(* IEC 61131-3 sources: SortJet_MasterSPS_Aufbau.fbsproj/07_Auftragsverwaltung/Job_Shuttle.prg.st^, 9 files *)

(* ---- Auftraege.act.st ---- *)
(* METADATA
{
	"v3Meta": {
		"objectGuid": "374beb49-ca7f-40e9-b2ab-7b5100759e7c"
	}
}
*)
ACTION Auftraege
//-------------------------------------------------------------------------------------------------
// AUFTRAG: M_SB0_MMI_SHEET_ORDER_SHUTTLE
//-------------------------------------------------------------------------------------------------
(* Hinweis:
   - Auftragsdaten an ein Shuttle uebergeben
*)
IF ( M_SB0_MMI_SHEET_ORDER_SHUTTLE ) THEN

  CASE tMmi2SpsInfo.wStationsNr OF

    cERSTES_SHUTTLE..cLETZTES_SHUTTLE:
      LocalAuftragsSpeicher REF= AuftragsSpeicherWand[tMmi2SpsInfo.wStationsNr, tMmi2SpsInfo.wAuftragsWand];
      M_SB0_MMI_SHEET_ORDER_SHUTTLE := FALSE;

    cERSTES_TRANSFERSHUTTLE..cLETZTES_TRANSFERSHUTTLE:
      LocalAuftragsSpeicher REF= AuftragsSpeicherTransfershuttle[tMmi2SpsInfo.wStationsNr];
      M_SB0_MMI_SHEET_ORDER_SHUTTLE := FALSE;

  END_CASE

  IF __ISVALIDREF(LocalAuftragsSpeicher) THEN

    LocalAuftragsSpeicher.NeuerAuftrag.wStationsNr            := tMmi2SpsInfo.wStationsNr;
    LocalAuftragsSpeicher.NeuerAuftrag.rVorabPosition         := tMmi2SpsInfo.rStationsPosition;
    LocalAuftragsSpeicher.NeuerAuftrag.rStationsZielposition  := tMmi2SpsInfo.rStationsPosition;     // Stationsposition der Quellstation
    LocalAuftragsSpeicher.NeuerAuftrag.rAuftragsLaenge        := tMmi2SpsInfo.rAuftragsLaenge;       // Länge der Scheibe/Batch
    LocalAuftragsSpeicher.NeuerAuftrag.rAuftragsHoehe         := tMmi2SpsInfo.rAuftragsHoehe;        // Höhe der Scheibe/Batch
    LocalAuftragsSpeicher.NeuerAuftrag.rAuftragsDicke         := tMmi2SpsInfo.rAuftragsDicke;        // Dicke der Scheibe/Batch
    LocalAuftragsSpeicher.NeuerAuftrag.wErsteLetzteScheibe    := tMmi2SpsInfo.wErsteLetzteScheibe;  // Kennzeichnung Erste und Letzte Scheibe
    LocalAuftragsSpeicher.NeuerAuftrag.wAnzahlScheiben        := tMmi2SpsInfo.wAnzahlScheiben;       // Anzahl der Scheiben
    LocalAuftragsSpeicher.NeuerAuftrag.wStationsWand          := tMmi2SpsInfo.wAuftragsWand;         // Stationswand der Quellstation
    LocalAuftragsSpeicher.NeuerAuftrag.wTransferstationsNr1   := tMmi2SpsInfo.wTransferstationsNr1;  // Stationsnummer der Zielstation 1
    LocalAuftragsSpeicher.NeuerAuftrag.wTransferstationsNr2   := tMmi2SpsInfo.wTransferstationsNr2;  // Stationsnummer der Zielstation 2
    LocalAuftragsSpeicher.NeuerAuftrag.rTransferposition1     := tMmi2SpsInfo.rTransferposition1;    // Stationsposition der Zielstation 1
    LocalAuftragsSpeicher.NeuerAuftrag.rTransferposition2     := tMmi2SpsInfo.rTransferposition2;    // Stationsposition der Zielstation 2
    LocalAuftragsSpeicher.NeuerAuftrag.wTransferwand          := tMmi2SpsInfo.wTransferwand;         // Stationswand der Zielstationen 1
    LocalAuftragsSpeicher.NeuerAuftrag.stAuftragsInformationen.wAuftragsInformationen := tMmi2SpsInfo.wAuftragsTyp;            // Zusaetzliche Auftrags- Informationen

    // Soll Drehpos der Folgestation für den Eintransport
    LocalAuftragsSpeicher.NeuerAuftrag.wTransferVersatzVorne   := tMmi2SpsInfo.rTransferstationModellversatzVorne;
    // Soll Drehpos der Folgestation nach dem Eintransport
    LocalAuftragsSpeicher.NeuerAuftrag.wTransferVersatzHinten  := tMmi2SpsInfo.rTransferstationModellversatzHinten;

    (* Hinweis:
       - Zuweisung der Bits "erste" und "letzte" Scheibe
    *)
    ErsteUndLetzteScheibeBits( wpErsteUndLetzteScheibe:= tMmi2SpsInfo.wErsteLetzteScheibe ,
                               wpLetzteScheibe => wlLetzteScheibe,
                               wpErsteScheibe  => wlErsteScheibe );

    LocalAuftragsSpeicher.NeuerAuftrag.bLetzteScheibe  := wlLetzteScheibe > 0;   // Stationsposition der Zielstation 2
    LocalAuftragsSpeicher.NeuerAuftrag.bErsteScheibe   := wlErsteScheibe  > 0;        // Stationswand der Zielstationen

    (* Hinweis:
       - 0 -> Eintransport
       - 1 -> Austransport
    *)
    IF ( tMmi2SpsInfo.wAuftragsTyp.0 ) THEN
      LocalAuftragsSpeicher.NeuerAuftrag.wAuftrag := eStation_Austransport;
    ELSE
      LocalAuftragsSpeicher.NeuerAuftrag.wAuftrag := eStation_Eintransport;
    END_IF

    LocalAuftragsSpeicher(bpNeuerAuftrag := TRUE);

  END_IF

END_IF

//-------------------------------------------------------------------------------------------------
// AUFTRAG: M_SB0_MMI_SortierungInsertExtractionShuttleData
//-------------------------------------------------------------------------------------------------
(* Hinweis:
   - Austransportschlitten mit einem Scheibenvortransport-Auftrag versehen
*)
IF ( M_SB0_MMI_SortierungInsertExtractionShuttleData ) THEN

  M_SB0_MMI_SortierungInsertExtractionShuttleData := FALSE;

  IF ( bgTransfershuttleVortransportAktivieren ) THEN

    // ---------------------------------------------------------------------------------------
    //  TRANSFERSHUTTLE VORTRANSPORT
    //
    //  Hinweis:
    //  - VortransportNummer_TS2 = 0   => Vortransport mit nur einem Transfershuttle
    //  - VortransportNummer_TS1 <> 0  => Vortransport im Transfershuttle-Verbund
    // ---------------------------------------------------------------------------------------
    IF ( tMmi2SpsInfo.wVortransportNummer_TS2 = 0  ) THEN

      AuftragsSpeicherTransfershuttle[tMmi2SpsInfo.wVortransportNummer_TS1].NeuerAuftrag.rStationsZielposition := tMmi2SpsInfo.rVortransportSollPosition_TS1;
      AuftragsSpeicherTransfershuttle[tMmi2SpsInfo.wVortransportNummer_TS1].NeuerAuftrag.rAuftragsLaenge       := tMmi2SpsInfo.rVortransportStrecke;
      AuftragsSpeicherTransfershuttle[tMmi2SpsInfo.wVortransportNummer_TS1].NeuerAuftrag.wTransferstationsNr1  := 0;
      AuftragsSpeicherTransfershuttle[tMmi2SpsInfo.wVortransportNummer_TS1].NeuerAuftrag.wTransferstationsNr2  := 0;
      AuftragsSpeicherTransfershuttle[tMmi2SpsInfo.wVortransportNummer_TS1].NeuerAuftrag.rTransferposition1    := tMmi2SpsInfo.rVortransportSollPosition_TS1;
      AuftragsSpeicherTransfershuttle[tMmi2SpsInfo.wVortransportNummer_TS1].NeuerAuftrag.rTransferposition2    := 0;
      AuftragsSpeicherTransfershuttle[tMmi2SpsInfo.wVortransportNummer_TS1].NeuerAuftrag.stAuftragsInformationen.cBIT_BUFFERSLOT_THICKNESS := ( tMmi2SpsInfo.wSlotThickness = 1 );
      AuftragsSpeicherTransfershuttle[tMmi2SpsInfo.wVortransportNummer_TS1].NeuerAuftrag.wAuftrag := eStation_Vortransport;
      AuftragsSpeicherTransfershuttle[tMmi2SpsInfo.wVortransportNummer_TS1](bpNeuerAuftrag := TRUE);

    ELSE
      VailiderenTransfershuttleVerbund ( wTransferstation1 := tMmi2SpsInfo.wVortransportNummer_TS1 ,
                                         wTransferstation2 := tMmi2SpsInfo.wVortransportNummer_TS2 ,
                                         wTransferstationMaster => tMmi2SpsInfo.wVortransportNummer_TS1,
                                         wTransferstationSlave  => tMmi2SpsInfo.wVortransportNummer_TS2 );

      AuftragsSpeicherTransfershuttle[tMmi2SpsInfo.wVortransportNummer_TS1].NeuerAuftrag.rStationsZielposition := tMmi2SpsInfo.rVortransportSollPosition_TS1;
      AuftragsSpeicherTransfershuttle[tMmi2SpsInfo.wVortransportNummer_TS1].NeuerAuftrag.rAuftragsLaenge       := tMmi2SpsInfo.rVortransportStrecke;
      AuftragsSpeicherTransfershuttle[tMmi2SpsInfo.wVortransportNummer_TS1].NeuerAuftrag.wTransferstationsNr1  := tMmi2SpsInfo.wVortransportNummer_TS1;
      AuftragsSpeicherTransfershuttle[tMmi2SpsInfo.wVortransportNummer_TS1].NeuerAuftrag.wTransferstationsNr2  := tMmi2SpsInfo.wVortransportNummer_TS2;
      AuftragsSpeicherTransfershuttle[tMmi2SpsInfo.wVortransportNummer_TS1].NeuerAuftrag.rTransferposition1    := tMmi2SpsInfo.rVortransportSollPosition_TS1;
      AuftragsSpeicherTransfershuttle[tMmi2SpsInfo.wVortransportNummer_TS1].NeuerAuftrag.rTransferposition2    := tMmi2SpsInfo.rVortransportSollPosition_TS2;
      AuftragsSpeicherTransfershuttle[tMmi2SpsInfo.wVortransportNummer_TS1].NeuerAuftrag.stAuftragsInformationen.cBIT_BUFFERSLOT_THICKNESS := ( tMmi2SpsInfo.wSlotThickness = 1 );
      AuftragsSpeicherTransfershuttle[tMmi2SpsInfo.wVortransportNummer_TS1].NeuerAuftrag.wAuftrag              := eStation_Vortransport;
      AuftragsSpeicherTransfershuttle[tMmi2SpsInfo.wVortransportNummer_TS1](bpNeuerAuftrag := TRUE);

    END_IF

  ELSE

    (* Hinweis:
       - Quittierung des Vortransportes
    *)
    wSps2MmiQuittierungVortransportStationsNr1 := tMmi2SpsInfo.wVortransportNummer_TS1;
    wSps2MmiQuittierungVortransportStationsNr2 := tMmi2SpsInfo.wVortransportNummer_TS2;
    wSps2MmiQuittierungVortransportStatus      := 1; // 0  = nicht Erfolgreich / 1 = erfolgreich
    rSps2MmiQuittierungVortransportWegStrecke  := tMmi2SpsInfo.rVortransportStrecke;

    MsgToMmi(auftragsnr_w := SB0_SPS_SortierungQuittExtractionShuttleData );

  END_IF

END_IF

//-------------------------------------------------------------------------------------------------
// AUFTRAG: M_SB0_MMI_SHUTTLE_INFORMATION
//-------------------------------------------------------------------------------------------------
IF ( M_SB0_MMI_SHUTTLE_INFORMATION ) THEN

  M_SB0_MMI_SHUTTLE_INFORMATION := FALSE;

  CASE tMmi2SpsInfo.wAuftrag_ShuttleNummer OF

    cERSTE_STATION..cLETZTE_STATION:
      ;
    cERSTES_SHUTTLE..cLETZTES_SHUTTLE:
      // Rueckfall: Schickt das MMI keine Wand (0), gilt Wand 1
      IF tMmi2SpsInfo.wAuftrag_ShuttleWand = 0 THEN
        tMmi2SpsInfo.wAuftrag_ShuttleWand := cWAND_1;
      END_IF
      CASE tMmi2SpsInfo.wAuftrag_ShuttleWand OF

          cWAND_1,
            cWAND_2:
          IF ( VorAbAuftragsDaten[tMmi2SpsInfo.wAuftrag_ShuttleNummer, tMmi2SpsInfo.wAuftrag_ShuttleWand].wAuftrag = eStation_Kein_Auftrag ) THEN
            VorAbAuftragsDaten[tMmi2SpsInfo.wAuftrag_ShuttleNummer, tMmi2SpsInfo.wAuftrag_ShuttleWand].rLaenge                := tMmi2SpsInfo.rAuftrag_Laenge;
            VorAbAuftragsDaten[tMmi2SpsInfo.wAuftrag_ShuttleNummer, tMmi2SpsInfo.wAuftrag_ShuttleWand].rDicke                 := tMmi2SpsInfo.rAuftrag_Dicke;
            VorAbAuftragsDaten[tMmi2SpsInfo.wAuftrag_ShuttleNummer, tMmi2SpsInfo.wAuftrag_ShuttleWand].wTransferStation       := tMmi2SpsInfo.wAuftrag_TranferStation;
            VorAbAuftragsDaten[tMmi2SpsInfo.wAuftrag_ShuttleNummer, tMmi2SpsInfo.wAuftrag_ShuttleWand].wAuftragstyp           := tMmi2SpsInfo.wAuftrag_Modus;
            VorAbAuftragsDaten[tMmi2SpsInfo.wAuftrag_ShuttleNummer, tMmi2SpsInfo.wAuftrag_ShuttleWand].wShuttleWandNummer     := tMmi2SpsInfo.wAuftrag_ShuttleWand;
            VorAbAuftragsDaten[tMmi2SpsInfo.wAuftrag_ShuttleNummer, tMmi2SpsInfo.wAuftrag_ShuttleWand].wTransferWand          := tMmi2SpsInfo.wAuftrag_TransferWand;
            VorAbAuftragsDaten[tMmi2SpsInfo.wAuftrag_ShuttleNummer, tMmi2SpsInfo.wAuftrag_ShuttleWand].wShuttleNummer         := tMmi2SpsInfo.wAuftrag_ShuttleNummer;

            VorAbAuftragsDaten[tMmi2SpsInfo.wAuftrag_ShuttleNummer, tMmi2SpsInfo.wAuftrag_ShuttleWand].stAuftragsInformationen.wAuftragsInformationen := tMmi2SpsInfo.wAuftrag_Modus;
            VorAbAuftragsDaten[tMmi2SpsInfo.wAuftrag_ShuttleNummer, tMmi2SpsInfo.wAuftrag_ShuttleWand].wAuftrag := eStation_VorabAuftrag;

          END_IF

        cWAND_1_2: //eigentlich Wand 1 und 2, da dies Bitcodiert ist, kommt dies als Wand3
          FOR wlIndexWand := cWAND_1 TO cANZAHL_WAENDE DO

            IF ( VorAbAuftragsDaten[tMmi2SpsInfo.wAuftrag_ShuttleNummer, wlIndexWand].wAuftrag = eStation_Kein_Auftrag ) THEN

              VorAbAuftragsDaten[tMmi2SpsInfo.wAuftrag_ShuttleNummer, wlIndexWand].rLaenge                := tMmi2SpsInfo.rAuftrag_Laenge;
              VorAbAuftragsDaten[tMmi2SpsInfo.wAuftrag_ShuttleNummer, wlIndexWand].rDicke                 := tMmi2SpsInfo.rAuftrag_Dicke;
              VorAbAuftragsDaten[tMmi2SpsInfo.wAuftrag_ShuttleNummer, wlIndexWand].wTransferStation       := tMmi2SpsInfo.wAuftrag_TranferStation;
              VorAbAuftragsDaten[tMmi2SpsInfo.wAuftrag_ShuttleNummer, wlIndexWand].wAuftragstyp           := tMmi2SpsInfo.wAuftrag_Modus;
              VorAbAuftragsDaten[tMmi2SpsInfo.wAuftrag_ShuttleNummer, wlIndexWand].wShuttleWandNummer     := wlIndexWand;
              VorAbAuftragsDaten[tMmi2SpsInfo.wAuftrag_ShuttleNummer, wlIndexWand].wTransferWand          := tMmi2SpsInfo.wAuftrag_TransferWand;
              VorAbAuftragsDaten[tMmi2SpsInfo.wAuftrag_ShuttleNummer, wlIndexWand].wShuttleNummer         := tMmi2SpsInfo.wAuftrag_ShuttleNummer;

              VorAbAuftragsDaten[tMmi2SpsInfo.wAuftrag_ShuttleNummer, wlIndexWand].stAuftragsInformationen.wAuftragsInformationen := tMmi2SpsInfo.wAuftrag_Modus;
              VorAbAuftragsDaten[tMmi2SpsInfo.wAuftrag_ShuttleNummer, wlIndexWand].wAuftrag := eStation_VorabAuftrag;

            END_IF

          END_FOR

        ELSE
          ;

      END_CASE

    cERSTES_TRANSFERSHUTTLE..cLETZTES_TRANSFERSHUTTLE:
      IF ( NOT Job_Shuttle.abpStarteParalleleBausteinAnsteuerung[tMmi2SpsInfo.wAuftrag_ShuttleNummer] ) THEN
        Job_Shuttle.VorAbAuftragsDaten[tMmi2SpsInfo.wAuftrag_ShuttleNummer, cWAND_1].rLaenge                := tMmi2SpsInfo.rAuftrag_Laenge;
        Job_Shuttle.VorAbAuftragsDaten[tMmi2SpsInfo.wAuftrag_ShuttleNummer, cWAND_1].rDicke                 := tMmi2SpsInfo.rAuftrag_Dicke;
        Job_Shuttle.VorAbAuftragsDaten[tMmi2SpsInfo.wAuftrag_ShuttleNummer, cWAND_1].wTransferStation       := tMmi2SpsInfo.wAuftrag_TranferStation;
        Job_Shuttle.VorAbAuftragsDaten[tMmi2SpsInfo.wAuftrag_ShuttleNummer, cWAND_1].wAuftragstyp           := tMmi2SpsInfo.wAuftrag_Modus;
        Job_Shuttle.VorAbAuftragsDaten[tMmi2SpsInfo.wAuftrag_ShuttleNummer, cWAND_1].wShuttleWandNummer     := tMmi2SpsInfo.wAuftrag_ShuttleWand;
        Job_Shuttle.VorAbAuftragsDaten[tMmi2SpsInfo.wAuftrag_ShuttleNummer, cWAND_1].wTransferWand          := tMmi2SpsInfo.wAuftrag_TransferWand;
        Job_Shuttle.VorAbAuftragsDaten[tMmi2SpsInfo.wAuftrag_ShuttleNummer, cWAND_1].wShuttleNummer         := tMmi2SpsInfo.wAuftrag_ShuttleNummer;

        Job_Shuttle.VorAbAuftragsDaten[tMmi2SpsInfo.wAuftrag_ShuttleNummer, cWAND_1].stAuftragsInformationen.wAuftragsInformationen := tMmi2SpsInfo.wAuftrag_Modus;

        Job_Shuttle.abpStarteParalleleBausteinAnsteuerung[tMmi2SpsInfo.wAuftrag_ShuttleNummer] := TRUE;
      END_IF

    ELSE
      (* Fehlerbehandlung:
      *)
      wpgFehlerdaten[0] := tMmi2SpsInfo.wAuftrag_ShuttleNummer;
      wpgFehlerdaten[1] := tMmi2SpsInfo.wAuftrag_TranferStation;
      SpsError( eFehler_Station,
                cMELDUNG_AUFTRAGSDATEN_UNGUELTIGE_STATION,
                tMmi2SpsInfo.wAuftrag_ShuttleNummer,
                AutomatikkreisBestimmen(tMmi2SpsInfo.wAuftrag_ShuttleNummer),
                wpgFehlerdaten );

  END_CASE

END_IF

//-------------------------------------------------------------------------------------------------
// AUFTRAG: M_SB0_MMI_GETSORTIERUNGSHUTTLEPOS
//-------------------------------------------------------------------------------------------------
(* Hinweis:
   - Verfarhlogik
     => Absetzen der Positionen
     => Melden der IST- Position wenn die Positionierung aufgrund eines
        Fehler [ Verfahrfreigabe fehlt ] nicht durchgefuehrt werden kann
*)
IF ( M_SB0_MMI_GETSORTIERUNGSHUTTLEPOS ) THEN

  M_SB0_MMI_GETSORTIERUNGSHUTTLEPOS := FALSE;

  SendShuttlePosition();

END_IF

//-------------------------------------------------------------------------------------------------
// AUFTRAG: M_SB0_MMI_TS_REPOSITIONING_LITES
//-------------------------------------------------------------------------------------------------

(* Hinweis:
   - Funktion zum zurueckfahren der Glaeser und neu Positionieren im Speicher
*)
IF ( M_SB0_MMI_TS_REPOSITIONING_LITES ) THEN
  M_SB0_MMI_TS_REPOSITIONING_LITES := FALSE;

  CASE tMmi2SpsInfo.wStationsNr OF

    cERSTES_TRANSFERSHUTTLE..cLETZTES_TRANSFERSHUTTLE:
      AuftragsSpeicherTransfershuttle[tMmi2SpsInfo.wStationsNr].NeuerAuftrag.wStationsNr           := tMmi2SpsInfo.wStationsNr;
      AuftragsSpeicherTransfershuttle[tMmi2SpsInfo.wStationsNr].NeuerAuftrag.rStationsZielposition := tMmi2SpsInfo.rStationsPosition;
      AuftragsSpeicherTransfershuttle[tMmi2SpsInfo.wStationsNr].NeuerAuftrag.wTransferstationsNr1  := tMmi2SpsInfo.wTransferstationsNr1;
      AuftragsSpeicherTransfershuttle[tMmi2SpsInfo.wStationsNr].NeuerAuftrag.rModellVersatzHinten  := tMmi2SpsInfo.rModellversatzHinten;

      IF ( tMmi2SpsInfo.rAuftragsDicke = 0 ) THEN
        AuftragsSpeicherTransfershuttle[tMmi2SpsInfo.wStationsNr].NeuerAuftrag.rAuftragsDicke        := 4.0;
      ELSE
        AuftragsSpeicherTransfershuttle[tMmi2SpsInfo.wStationsNr].NeuerAuftrag.rAuftragsDicke        := 19.0;
      END_IF

      AuftragsSpeicherTransfershuttle[tMmi2SpsInfo.wStationsNr].NeuerAuftrag.wAuftrag := eStation_Scheibenkorrektur;
      AuftragsSpeicherTransfershuttle[tMmi2SpsInfo.wStationsNr](bpNeuerAuftrag := TRUE);

      AuftragsSpeicherTransfershuttle[tMmi2SpsInfo.wTransferstationsNr1].NeuerAuftrag.wStationsNr           := tMmi2SpsInfo.wTransferstationsNr1;
      AuftragsSpeicherTransfershuttle[tMmi2SpsInfo.wTransferstationsNr1].NeuerAuftrag.rStationsZielposition := tMmi2SpsInfo.rTransferposition1;
      AuftragsSpeicherTransfershuttle[tMmi2SpsInfo.wTransferstationsNr1].NeuerAuftrag.wTransferstationsNr1  := tMmi2SpsInfo.wStationsNr;
      AuftragsSpeicherTransfershuttle[tMmi2SpsInfo.wTransferstationsNr1].NeuerAuftrag.rModellVersatzHinten  := tMmi2SpsInfo.rModellversatzHinten;

      IF ( tMmi2SpsInfo.rAuftragsDicke = 0 ) THEN
        AuftragsSpeicherTransfershuttle[tMmi2SpsInfo.wTransferstationsNr1].NeuerAuftrag.rAuftragsDicke        := 4.0;
      ELSE
        AuftragsSpeicherTransfershuttle[tMmi2SpsInfo.wTransferstationsNr1].NeuerAuftrag.rAuftragsDicke        := 19.0;
      END_IF

      AuftragsSpeicherTransfershuttle[tMmi2SpsInfo.wTransferstationsNr1].NeuerAuftrag.wAuftrag := eStation_Transportkopplung;
      AuftragsSpeicherTransfershuttle[tMmi2SpsInfo.wTransferstationsNr1](bpNeuerAuftrag := TRUE);

  END_CASE

END_IF

//-------------------------------------------------------------------------------------------------
// AUFTRAG: M_SB0_MMI_SORTIERUNGCANcELSHUTTLEDATA
//-------------------------------------------------------------------------------------------------
(* Hinweis:
   - Abbrechen eines aktiven Shuttleauftrags
*)
IF ( M_SB0_MMI_SORTIERUNGCANCELSHUTTLEDATA ) THEN

  M_SB0_MMI_SortierungCancelShuttleData := FALSE;

  CASE tMmi2SpsInfo.wCancelShuttleDataShuttleNr OF

    cERSTES_SHUTTLE..cLETZTES_SHUTTLE:
      IF ( AuftragsdatenWand[tMmi2SpsInfo.wCancelShuttleDataShuttleNr, cWAND_1].wAuftrag <> eStation_Kein_Auftrag ) THEN
        AuftragsdatenWand[tMmi2SpsInfo.wCancelShuttleDataShuttleNr, cWAND_1].wAuftrag :=  eStation_Kein_Auftrag;
      END_IF

    cERSTES_TRANSFERSHUTTLE..cLETZTES_TRANSFERSHUTTLE:
      IF ( Job_Shuttle.AuftragsdatenTransfershuttle[tMmi2SpsInfo.wCancelShuttleDataShuttleNr].wAuftrag <> eStation_Kein_Auftrag ) THEN
        Job_Shuttle.AuftragsdatenTransfershuttle[tMmi2SpsInfo.wCancelShuttleDataShuttleNr].wAuftrag :=  eStation_Kein_Auftrag;
      END_IF

  END_CASE

END_IF

//-------------------------------------------------------------------------------------------------
// S T A R T - Fächerwagen Suche mittels Sensor
//-------------------------------------------------------------------------------------------------

IF ( M_SB0_MMI_POSITIONMEASUREONOFF ) THEN

  M_SB0_MMI_POSITIONMEASUREONOFF := FALSE;

  IF ( tMmi2SpsInfo.wShuttleFWSucheAN_AUS = 1 ) THEN
    AuftragsSpeicherWand[tMmi2SpsInfo.wShuttleNummerFWSuche, cWAND_1].NeuerAuftrag.wAuftrag := eStation_RackSuche;
    AuftragsSpeicherWand[tMmi2SpsInfo.wShuttleNummerFWSuche, cWAND_1](bpNeuerAuftrag := TRUE);
  ELSE
    IF ( AuftragsdatenWand[tMmi2SpsInfo.wShuttleNummerFWSuche, cWAND_1].wAuftrag = eStation_RackSuche ) THEN
      AuftragsdatenWand[tMmi2SpsInfo.wShuttleNummerFWSuche, cWAND_1].wAuftrag := eStation_Kein_Auftrag;
    END_IF
  END_IF

END_IF

//-------------------------------------------------------------------------------------------------
// SHUTTLE DEAKTIVIEREN VIA MMI
//-------------------------------------------------------------------------------------------------
IF ( M_SB0_MMI_STATIONSTATUS ) THEN

  CASE tMmi2SpsInfo.wStationsNummer OF

    cERSTES_SHUTTLE..cLETZTES_SHUTTLE:
      starrShuttleBasisParameter[tMmi2SpsInfo.wStationsNummer].stMKs.bDeaktivieren := tMmi2SpsInfo.wStationsStatusWord2.0;
      M_SB0_MMI_STATIONSTATUS := FALSE;

    cERSTES_TRANSFERSHUTTLE..cLETZTES_TRANSFERSHUTTLE:
      starrTransfershuttleBasisParameter[tMmi2SpsInfo.wStationsNummer].stMKs.bDeaktivieren := tMmi2SpsInfo.wStationsStatusWord2.0;
      M_SB0_MMI_STATIONSTATUS := FALSE;

  END_CASE

END_IF
END_ACTION

(* ---- Master_Transfershuttle.meth.st ---- *)
(* METADATA
{
	"v3Meta": {
		"objectGuid": "5a2b5255-704a-40f5-acbe-9caa573edc30"
	}
}
*)
METHOD INTERNAL Master_Transfershuttle
VAR_INPUT
  wStation : WORD;
END_VAR

// ****************************************************9*********************************************
// STEUERUNG: EINTRANSPORT
// *************************************************************************************************

IF ( AuftragsdatenTransfershuttle[wStation].wAuftrag = eStation_Eintransport ) THEN
  (* Hinweis:
     - Aufruf der Schrittkette
  *)
  TS_Eintransport[wStation]( Auftragsdaten := AuftragsdatenTransfershuttle[wStation], wStation := wStation );
  (* Hinweis:
     - Abschluss der Schrittkette
  *)
  IF TS_Eintransport[wStation].bpDone THEN
    AuftragsdatenTransfershuttle[wStation] := TS_Eintransport[wStation].Auftragsdaten;
    TS_Eintransport[wStation](bpReset := TRUE);
  END_IF
  (* Hinweis:
     - Fehler-Auswertung
  *)
  blFehlerTS[wStation] := TS_Eintransport[wStation].bpFehler;
  IF rtlFehlerTS[wStation].Q THEN
    IF ( starrTransfershuttleBasisParameter[wStation].bRueckwaertsTransportieren[cWAND_1] ) THEN
      AutomatikFehlerTransfershuttleSetzen(starrTransferShuttleBasisParameter[wStation].stMKs.eaAutomatikkreis, abpFehler, cSPEICHER_AUSLAUFSEITE);
      IF aTransfershuttles[wStation].bpAnforderungBetriebsstopp THEN
        AutomatikFehlerTransfershuttleSetzen(starrTransferShuttleBasisParameter[wStation].stMKs.eaAutomatikkreis, abpFehler, cSPEICHER_EINLAUFSEITE);
      END_IF
    ELSE
      AutomatikFehlerTransfershuttleSetzen(starrTransferShuttleBasisParameter[wStation].stMKs.eaAutomatikkreis, abpFehler, cSPEICHER_EINLAUFSEITE);
      IF aTransfershuttles[wStation].bpAnforderungBetriebsstopp THEN
        AutomatikFehlerTransfershuttleSetzen(starrTransferShuttleBasisParameter[wStation].stMKs.eaAutomatikkreis, abpFehler, cSPEICHER_AUSLAUFSEITE);
      END_IF
    END_IF
  END_IF
ELSE
  (* Hinweis:
     - Reset der Schrittkette
  *)
  IF ( TS_Eintransport[wStation].steplSchritt <> STEP_0_E ) THEN
    TS_Eintransport[wStation](bpReset := TRUE);
  END_IF
END_IF

// ****************************************************9*********************************************
// STEUERUNG: AUSTRANSPORT
// *************************************************************************************************

IF ( AuftragsdatenTransfershuttle[wStation].wAuftrag = eStation_Austransport ) THEN
  (* Hinweis:
     - Aufruf der Schrittkette
  *)
  TS_Austransport[wStation]( Auftragsdaten := AuftragsdatenTransfershuttle[wStation], wStation := wStation );
  (* Hinweis:
     - Abschluss der Schrittkette
  *)
  IF TS_Austransport[wStation].bpDone THEN
    AuftragsdatenTransfershuttle[wStation] := TS_Austransport[wStation].Auftragsdaten;
    TS_Austransport[wStation](bpReset := TRUE);
  END_IF
  (* Hinweis:
     - Fehler-Auswertung
  *)
  blFehlerTS[wStation] := TS_Austransport[wStation].bpFehler;
  IF rtlFehlerTS[wStation].Q THEN
    IF ( starrTransfershuttleBasisParameter[wStation].bRueckwaertsTransportieren[cWAND_1] ) THEN
      AutomatikFehlerTransfershuttleSetzen(starrTransferShuttleBasisParameter[wStation].stMKs.eaAutomatikkreis, abpFehler, cSPEICHER_EINLAUFSEITE);
      IF aTransfershuttles[wStation].bpAnforderungBetriebsstopp THEN
        AutomatikFehlerTransfershuttleSetzen(starrTransferShuttleBasisParameter[wStation].stMKs.eaAutomatikkreis, abpFehler, cSPEICHER_AUSLAUFSEITE);
      END_IF
    ELSE
      AutomatikFehlerTransfershuttleSetzen(starrTransferShuttleBasisParameter[wStation].stMKs.eaAutomatikkreis, abpFehler, cSPEICHER_AUSLAUFSEITE);
      IF aTransfershuttles[wStation].bpAnforderungBetriebsstopp THEN
        AutomatikFehlerTransfershuttleSetzen(starrTransferShuttleBasisParameter[wStation].stMKs.eaAutomatikkreis, abpFehler, cSPEICHER_EINLAUFSEITE);
      END_IF
    END_IF
  END_IF
ELSE
  (* Hinweis:
     - Reset der Schrittkette
  *)
  IF ( TS_Austransport[wStation].steplSchritt <> STEP_0_E ) THEN
    TS_Austransport[wStation](bpReset := TRUE);
  END_IF
END_IF

// ****************************************************9*********************************************
// STEUERUNG: VORTRANSPORT
// *************************************************************************************************

IF ( AuftragsdatenTransfershuttle[wStation].wAuftrag = eStation_Vortransport ) THEN
  (* Hinweis:
     - Aufruf der Schrittkette
  *)
  TS_Vortransport[wStation]( Auftragsdaten := AuftragsdatenTransfershuttle[wStation], wStation := wStation);
  (* Hinweis:
     - Abschluss der Schrittkette
  *)
  IF TS_Vortransport[wStation].bpDone THEN
    AuftragsdatenTransfershuttle[wStation] := TS_Vortransport[wStation].Auftragsdaten;
    TS_Vortransport[wStation](bpReset := TRUE);
  END_IF
  (* Hinweis:
     - Fehler-Auswertung
  *)
  blFehlerTS[wStation] := TS_Vortransport[wStation].bpFehler;
  IF rtlFehlerTS[wStation].Q THEN
    AutomatikFehlerSetzen(starrTransferShuttleBasisParameter[wStation].stMKs.eaAutomatikkreis, abpFehler);
  END_IF
ELSE
  (* Hinweis:
     - Reset der Schrittkette
  *)
  IF ( TS_Vortransport[wStation].steplSchritt <> STEP_0_E ) THEN
    TS_Vortransport[wStation](bpReset := TRUE);
  END_IF
END_IF

// ****************************************************9*********************************************
// STEUERUNG: QUERFAHRT
// *************************************************************************************************

IF ( AuftragsdatenTransfershuttle[wStation].wAuftrag = eStation_Vorabpositionierung ) THEN
  (* Hinweis:
     - Aufruf der Schrittkette
  *)
  TS_Querfahrt[wStation]( Auftragsdaten := AuftragsdatenTransfershuttle[wStation], wStation := wStation );
  (* Hinweis:
     - Abschluss der Schrittkette
  *)
  IF TS_Querfahrt[wStation].bpDone THEN
    AuftragsdatenTransfershuttle[wStation] := TS_Querfahrt[wStation].Auftragsdaten;
    TS_Querfahrt[wStation](bpReset := TRUE);
  END_IF
  (* Hinweis:
     - Fehler-Auswertung
  *)
  blFehlerTS[wStation] := TS_Querfahrt[wStation].bpFehler;
  IF rtlFehlerTS[wStation].Q THEN
    AutomatikFehlerSetzen(starrTransferShuttleBasisParameter[wStation].stMKs.eaAutomatikkreis, abpFehler);
  END_IF
ELSE
  (* Hinweis:
     - Reset der Schrittkette
  *)
  IF ( TS_Querfahrt[wStation].steplSchritt <> STEP_0_E ) THEN
    TS_Querfahrt[wStation](bpReset := TRUE);
  END_IF
END_IF

//-------------------------------------------------------------------------------------------------
// STEUERUNG: SPEICHERFACHVALIDIERUNG
//-------------------------------------------------------------------------------------------------
IF (  abpSpeicherfachValidierung[wStation] ) THEN
  CASE asteplSpeicherfachValidierung[wStation] OF
    // SPEICHERFACHVALIDIERUNG =============================
    STEP_0_E:
      (* Hinweis:
         - Option: Sicherstellen das der Output-Sicherheitskreis geschlossen ist
      *)
      IF checkSafetyCircuitsNotBlocked(starrTransferShuttleBasisParameter[wStation])
         AND NOT starrTransfershuttleBasisParameter[wStation].bReset
      THEN
        awlStatusSpeichervalidierung[wStation]   := cAUFTRAG_KEIN_STATUS;
        asteplSpeicherfachValidierung[wStation] := STEP_10_E;
      END_IF

    // SPEICHERFACHVALIDIERUNG =============================
    STEP_10_E:
      // ---------------------------------------------------------------------------------------
      //  PRUEFEN TRANSFERSHUTTLE VERBUND
      //
      //  Hinweis:
      //  - wTransfershuttle_Nummer2 = 0   => Vortransport mit nur einem Transfershuttle
      //  - wTransfershuttle_Nummer2 <> 0  => Vortransport im Transfershuttle-Verbund
      // ---------------------------------------------------------------------------------------

      IF ( starrAuftragsdatenSpeicherfachValidierung[wStation].wTransferstationsNr2 <> 0 )  THEN

        awlVerbundTransfershuttle[wStation] := AuftragsdatenTransfershuttle[wStation].wTransferstationsNr2;

        IF ( AuftragsdatenTransfershuttle[awlVerbundTransfershuttle[wStation]].wAuftrag = eStation_Kein_Auftrag ) THEN
          asteplSpeicherfachValidierung[wStation] := STEP_20_E;
        END_IF

      ELSE
        (* Hinweis:
           - Informationen uebergeben und die Validierung starten
        *)
        starrTransfershuttleBasisParameter[wStation].pAuftrag[cWAND_1] := starrAuftragsdatenSpeicherfachValidierung[wStation];
        aTransfershuttles[wStation].bpStarteSpeicherfachValidierung := TRUE;

        asteplSpeicherfachValidierung[wStation] := STEP_100_E;

      END_IF

    // SPEICHERFACHVALIDIERUNG =============================
    STEP_20_E:

      (* Hinweis:
         - Transfershuttle koppeln
      *)
      aTransfershuttles[wStation].stpInTransportVerbund                             := aTransfershuttles[awlVerbundTransfershuttle[wStation]].stpOutTransportVerbund;
      aTransfershuttles[awlVerbundTransfershuttle[wStation]].stpInTransportVerbund  := aTransfershuttles[wStation].stpOutTransportVerbund;

      (* Hinweis:
         - Auftragsdaten uebergeben
      *)
      AuftragsdatenTransfershuttle[awlVerbundTransfershuttle[wStation]].rAuftragsDicke        := starrAuftragsdatenSpeicherfachValidierung[wStation].rAuftragsDicke ;
      AuftragsdatenTransfershuttle[awlVerbundTransfershuttle[wStation]].rStationsZielposition := starrAuftragsdatenSpeicherfachValidierung[wStation].rTransferposition2 ;
      AuftragsdatenTransfershuttle[awlVerbundTransfershuttle[wStation]].wStationsNr           := starrAuftragsdatenSpeicherfachValidierung[wStation].wTransferstationsNr2 ;
      AuftragsdatenTransfershuttle[awlVerbundTransfershuttle[wStation]].wAuftrag              := eStation_Transportkopplung;

      (* Hinweis:
         - Auftragsdaten uebergeben
      *)
      starrTransfershuttleBasisParameter[wStation].pAuftrag[cWAND_1] := starrAuftragsdatenSpeicherfachValidierung[wStation];
      aTransfershuttles[wStation].bpStarteSpeicherfachValidierung := TRUE;

      asteplSpeicherfachValidierung[wStation] := STEP_100_E;

    // SPEICHERFACHVALIDIERUNG =============================
    STEP_100_E:
      // ---------------------------------------------------------------------------------------
      //  AUSWERTUNG TRANSFERSHUTTLE - SPEICHERFACH VALIDIERUNG
      //
      //  Hinweis:
      //  - n/c
      // ---------------------------------------------------------------------------------------

      IF ( aTransfershuttles[wStation].bpSpeicherfachValidierungAbgeschlossen ) THEN
        aTransfershuttles[wStation].bpStarteSpeicherfachValidierung := FALSE;
        awlStatusSpeichervalidierung[wStation] := cAUFTRAG_ERFOLGREICH;

        asteplSpeicherfachValidierung[wStation] := STEP_120_E;
      END_IF

      // Fehlverhalten
      IF ( starrTransfershuttleBasisParameter[wStation].bFehler ) THEN

        aTransfershuttles[wStation].bpStarteSpeicherfachValidierung := FALSE;
        awlStatusSpeichervalidierung[wStation] := cAUFTRAG_FEHLER;

        asteplSpeicherfachValidierung[wStation] := STEP_120_E;

        (* Hinweis:
           - Meldung an die HMI generieren.
             => Gesendet wird: Shuttlenummer \Position \Fehlertyp
        *)
        wgSps2MmiShuttleNr                 := starrTransfershuttleBasisParameter[wStation].stMKs.stStationsNummern.NummerIntern;
        rgSPS2MMIExtractionShuttlePosition := starrTransfershuttleBasisParameter[wStation].rAktuellePositionQuerfahrt;
        wSps2MmiFehlertyp                  := aTransfershuttles[wStation].wpAusnahmefehlerTyp;
        MsgToMmi(auftragsnr_w := SB0_SPS_TRANSFERSHUTTLEFEHLER );// Fehlermeldung ans MMI für den folgenden Systemcheck

        (* Hinweis:
           - Fehlermeldung generieren
        *)
        SpsError( eFehler_Station,
                  starrTransfershuttleBasisParameter[wStation].wFehlerNummer,
                  starrTransfershuttleBasisParameter[wStation].stMKs.stStationsNummern.NummerIntern,
                  AutomatikkreisBestimmen(starrTransfershuttleBasisParameter[wStation].stMKs.stStationsNummern.NummerSPS),
                  starrTransfershuttleBasisParameter[wStation].awFehlerInformationen );

      END_IF

    // SPEICHERFACHVALIDIERUNG =============================
    STEP_120_E:
      wgSps2MmiShuttleNr         := starrTransfershuttleBasisParameter[wStation].stMKs.stStationsNummern.NummerIntern;
      wSps2MmiValidierungsStatus := awlStatusSpeichervalidierung[wStation];
      MsgToMmi(auftragsnr_w := SB0_SPS_TRANSFERSHUTTLECHECK_ABGESCHLOSSEN );// Fehlermeldung ans MMI für den folgenden Systemcheck

      asteplSpeicherfachValidierung[wStation] := SEL( awlStatusSpeichervalidierung[wStation] = cAUFTRAG_FEHLER,
                                                      STEP_1000_E,
                                                      STEP_900_E );

    // SPEICHERFACHVALIDIERUNG =============================
    STEP_900_E:
      AutomatikFehlerSetzen(starrTransferShuttleBasisParameter[wStation].stMKs.eaAutomatikkreis, abpFehler);

    // SPEICHERFACHVALIDIERUNG =============================
    STEP_1000_E:
      abpSpeicherfachValidierung[wStation] := FALSE;

      (* Hinweis:
         - Pruefen ob die Transferkopplung geloest werden muss
      *)
      IF ( PruefungWertImIntervall(AuftragsdatenTransfershuttle[wStation].wTransferstationsNr2, cERSTES_TRANSFERSHUTTLE, cLETZTES_TRANSFERSHUTTLE) ) THEN

        IF ( AuftragsdatenTransfershuttle[AuftragsdatenTransfershuttle[wStation].wTransferstationsNr2].wAuftrag = eStation_Transportkopplung ) THEN
          AuftragsdatenTransfershuttle[AuftragsdatenTransfershuttle[wStation].wTransferstationsNr2].wAuftrag := eStation_Kein_Auftrag;
        END_IF

      END_IF

  // SPEICHERFACHVALIDIERUNG =============================
  END_CASE

END_IF

IF ( NOT abpSpeicherfachValidierung[wStation] ) THEN

  IF ( asteplSpeicherfachValidierung[wStation] > STEP_0_E ) THEN
    aTransfershuttles[wStation].bpStarteSpeicherfachValidierung := FALSE;
    asteplSpeicherfachValidierung[wStation] := STEP_0_E;
  END_IF

END_IF
END_METHOD

(* ---- Meldungen.act.st ---- *)
(* METADATA
{
	"v3Meta": {
		"objectGuid": "68e675d5-67ba-4597-82c1-c0511fb282bc"
	}
}
*)
ACTION Meldungen
//-------------------------------------------------------------------------------------------------
// AKTION: MELDUNGEN
//-------------------------------------------------------------------------------------------------
// WatchIO:
//   - Ueberwachung der Verfahrfreigabe der Shuttle
//     -> Inputshuttle
//     -> Outputshuttle
//     -> Transfershuttle
FOR wlIndex := cERSTES_SHUTTLE TO cLETZTES_SHUTTLE DO
  WatchIo( NOT abgVerfahrfreigabeShuttle[wlIndex], ioccShuttle1VerfahrfreigabeFehlt + (wlIndex - 101) );
END_FOR;

FOR wlIndex := cERSTES_TRANSFERSHUTTLE TO cLETZTES_TRANSFERSHUTTLE DO
  WatchIo( NOT abgVerfahrfreigabeShuttle[wlIndex], ioccTransfershuttle1VerfahrfreigabeFehlt + (wlIndex - 151) );
END_FOR;
END_ACTION

(* ---- Reset.act.st ---- *)
(* METADATA
{
	"v3Meta": {
		"objectGuid": "238ec719-f16e-4d9c-9f71-7a8241f71645"
	}
}
*)
ACTION Reset
//-------------------------------------------------------------------------------------------------
// AKTION: RESET
//-------------------------------------------------------------------------------------------------

(* Hinweis:
   - Zuruecksetzen des AK
     => Inputshuttle [expliziet]
*)
FOR wlIndexReset := cERSTER_AUTOMATIKKREIS TO cLETZTER_AUTOMATIKKREIS DO

  IF abpReset[wlIndexReset] THEN

    abpReset[wlIndexReset] := FALSE;
    abpFehler[wlIndexReset] := FALSE;

    FOR wlIndex := cERSTES_SHUTTLE TO cLETZTES_SHUTTLE DO
      IF StationInAutomatikkreis(starrShuttleBasisParameter[wlIndex].stMKs.eaAutomatikkreis, wlIndexReset) THEN
        AuftragsSpeicherShuttle[wlIndex].bpReset := TRUE;
        AuftragsSpeicherShuttle[wlIndex]();

        abgVerfahrfreigabeShuttle[wlindex] := TRUE;

        AuftragsdatenStation[wlIndex].wAuftrag := eStation_Kein_Auftrag;

        starrShuttleBasisParameter[wlIndex].bReset := TRUE;

        Querfahrt[wlIndex]( bpReset := TRUE );
        Racksuche[wlIndex]( bpReset := TRUE );

        FOR wlIndexWand := cWAND_1 TO cANZAHL_WAENDE DO

          AuftragsSpeicherWand[wlIndex,wlIndexWand].bpReset := TRUE;
          AuftragsSpeicherWand[wlIndex,wlIndexWand]();

          Eintransport[wlIndex, wlIndexWand]( bpReset := TRUE );
          Austransport[wlIndex, wlIndexWand]( bpReset := TRUE );

          VorabkomponentenAnsteuerung[wlIndex, wlIndexWand]( bpReset := TRUE );

          AuftragsdatenWand[wlIndex, wlIndexWand].wAuftrag := eStation_Kein_Auftrag;
          VorAbAuftragsDaten[wlIndex, wlIndexWand].wAuftrag := eStation_Kein_Auftrag;

          blFehler[wlIndex, wlIndexWand] := FALSE;

          starrShuttleBasisParameter[wlIndex].bEintransportGewesen[wlIndexWand] := FALSE;
        END_FOR

      END_IF
    END_FOR

    FOR wlIndex := cERSTES_TRANSFERSHUTTLE TO cLETZTES_TRANSFERSHUTTLE  DO

      // WICHTIG: OR_ELSE -> ZWEITE BEDINGUNG WIRD NUR GEPRÜFT, WENN ERSTE FALSE IST !!! IST DIE ERSTE FALSE, WIRD DIE 2. BEDINGUNG GEPRÜFT ; IST DIE ERSTE TRUE, WIRD DIE 2. BEDINGUNG IGNORIERT UND NICHT MEHR GEPRÜFT (wg. ZUGRIFFSVERLETZTUNG)
      // Alle konfigurierten Automatikkreise des TS sind in Hand
      // ODER
      // Output-AK ist nicht in den vorhandenen Automatikkreisen der Maschine definiert ; das heißt, Erster AK = 1 und ANZAHL < wlAutomatikkreis2 --- OR_ELSE der 2. konfigurierte Automatikkreis für das TS ist 0; somit ist das TS nur in einem AK definiert
      IF   ( NOT AutomatikAktiv(wlIndex)
             OR ( ( cANZAHL_AUTOMATIKKREISE = 1 ) OR_ELSE ( starrTransfershuttleBasisParameter[wlIndex].stMKs.eaAutomatikkreis[wlAutomatikkreis2] = 0 ) ) )
           AND StationInAutomatikkreis(starrTransfershuttleBasisParameter[wlIndex].stMKs.eaAutomatikkreis, wlIndexReset)
      THEN
        AuftragsSpeicherTransfershuttle[wlIndex].bpReset := TRUE;
        AuftragsSpeicherTransfershuttle[wlIndex]();

        abgVerfahrfreigabeShuttle[wlindex] := TRUE;

        abpStarteParalleleBausteinAnsteuerung[wlIndex] := FALSE;
        abpSpeicherfachValidierung[wlIndex]  := FALSE;
        AuftragsdatenTransfershuttle[wlIndex].wAuftrag := eStation_Kein_Auftrag;
        starrTransferShuttleBasisParameter[wlIndex].bReset := TRUE;
        blFehlerTS[wlIndex] := FALSE;

      ELSE

        // Der zu resettende AK entspricht dem ERSTEN (INPUTSEITE) konfigurierten AK des TS
        // UND Doppelte Sicherheit: Nochmal prüfen, dass das TS im zu resetten AK ist
        // UND Automatik des zu resettenden AK darf NICHT mehr TRUE sein
        IF                ( wlIndexReset = starrTransfershuttleBasisParameter[wlIndex].stMKs.eaAutomatikkreis[1] )
                 AND_THEN StationInAutomatikkreis(starrTransfershuttleBasisParameter[wlIndex].stMKs.eaAutomatikkreis, wlIndexReset)
                 AND_THEN NOT M_Automatik_Aktiv[starrTransfershuttleBasisParameter[wlIndex].stMKs.eaAutomatikkreis[1]]
        THEN
          IF ( ( ( AuftragsdatenTransfershuttle[wlIndex].wAuftrag = eStation_Eintransport )
                 OR ( AuftragsdatenTransfershuttle[wlIndex].wAuftrag = eStation_Scheibenkorrektur )
                 OR ( aTransfershuttles[wlIndex].ReservierungsStatus = TS_EINTRANSPORT_RESERVIERUNG )
                 OR ( aTransfershuttles[wlIndex].ReservierungsStatus = TS_AUSTRANSPORT_RUECKWERTIG_RESERVIERUNG ) )
               AND NOT aTransfershuttles[wlIndex].bpAnforderungBetriebsstopp )
          THEN
            AuftragsSpeicherTransfershuttle[wlIndex].bpReset := TRUE;
            AuftragsSpeicherTransfershuttle[wlIndex]();

            abgVerfahrfreigabeShuttle[wlindex] := TRUE;

            abpStarteParalleleBausteinAnsteuerung[wlIndex] := FALSE;
            abpSpeicherfachValidierung[wlIndex]  := FALSE;
            AuftragsdatenTransfershuttle[wlIndex].wAuftrag := eStation_Kein_Auftrag;
            starrTransferShuttleBasisParameter[wlIndex].bReset := TRUE;
            blFehlerTS[wlIndex] := FALSE;

            (* Hinweis:
               - Gilt nur fuer Systeme mit Master - Slave  Transfershuttle
            *)
            IF ( wlIndex MOD 2 = 1 ) AND ( UPPER_BOUND(AuftragsdatenTransfershuttle, 1 ) >= (wlIndex + 1) ) AND_THEN ( AuftragsdatenTransfershuttle[wlIndex + 1].wAuftrag = eStation_Transportkopplung ) THEN
              AuftragsdatenTransfershuttle[wlIndex + 1].wAuftrag := eStation_Kein_Auftrag;
              starrTransferShuttleBasisParameter[wlIndex + 1].bReset := TRUE;
            END_IF
          END_IF
        END_IF
        // Der zu resettende AK entspricht dem ZWEITEN (OUTPUTSEITE) konfigurierten AK des TS
        // WICHTIG: Erst pruefen, ob es ueberhaupt einen 2. AK gibt (Zugriffsverletzung bei nur einem AK)
        // UND Doppelte Sicherheit: Nochmal prüfen, dass das TS im zu resetten AK ist
        // UND Automatik des zu resettenden AK darf NICHT mehr TRUE sein
        IF                ( cANZAHL_AUTOMATIKKREISE > 1 )
                 AND_THEN ( starrTransfershuttleBasisParameter[wlIndex].stMKs.eaAutomatikkreis[wlAutomatikkreis2] <> 0 )
                 AND_THEN ( wlIndexReset =starrTransfershuttleBasisParameter[wlIndex].stMKs.eaAutomatikkreis[wlAutomatikkreis2] )
                 AND_THEN StationInAutomatikkreis(starrTransfershuttleBasisParameter[wlIndex].stMKs.eaAutomatikkreis, wlIndexReset)
                 AND_THEN NOT M_Automatik_Aktiv[starrTransfershuttleBasisParameter[wlIndex].stMKs.eaAutomatikkreis[wlAutomatikkreis2]]
        THEN
          IF ( ( ( AuftragsdatenTransfershuttle[wlIndex].wAuftrag = eStation_Austransport )
                 OR ( AuftragsdatenTransfershuttle[wlIndex].wAuftrag = eStation_Scheibenkorrektur )
                 OR ( aTransfershuttles[wlIndex].ReservierungsStatus = TS_AUSTRANSPORT_RESERVIERUNG )
                 OR ( aTransfershuttles[wlIndex].ReservierungsStatus = TS_EINTRANSPORT_RUECKWERTIG_RESERVIERUNG ) )
               AND NOT aTransfershuttles[wlIndex].bpAnforderungBetriebsstopp )
          THEN
            AuftragsSpeicherTransfershuttle[wlIndex].bpReset := TRUE;
            AuftragsSpeicherTransfershuttle[wlIndex]();

            abgVerfahrfreigabeShuttle[wlindex] := TRUE;

            abpStarteParalleleBausteinAnsteuerung[wlIndex] := FALSE;
            abpSpeicherfachValidierung[wlIndex]  := FALSE;
            AuftragsdatenTransfershuttle[wlIndex].wAuftrag := eStation_Kein_Auftrag;
            starrTransferShuttleBasisParameter[wlIndex].bReset := TRUE;
            blFehlerTS[wlIndex] := FALSE;
            (* Wichtig:
               - Gilt nur fuer Systeme mit Master - Slave  Transfershuttle-Verbund
            *)
            IF ( wlIndex MOD 2 = 1 ) AND ( UPPER_BOUND(AuftragsdatenTransfershuttle, 1 ) >= (wlIndex + 1) ) AND_THEN ( AuftragsdatenTransfershuttle[wlIndex + 1].wAuftrag = eStation_Transportkopplung ) THEN
              AuftragsdatenTransfershuttle[wlIndex + 1].wAuftrag := eStation_Kein_Auftrag;
              starrTransferShuttleBasisParameter[wlIndex + 1].bReset := TRUE;
            END_IF
          END_IF
        END_IF

      END_IF

    END_FOR

  END_IF

END_FOR
END_ACTION

(* ---- ShuttleQuerfahrt.meth.st ---- *)
(* METADATA
{
	"v3Meta": {
		"objectGuid": "c062f55a-4f6a-45c2-9de2-37ec00cd7b53"
	}
}
*)
METHOD INTERNAL ShuttleQuerfahrt
VAR_INPUT
  wStation : WORD;
END_VAR

// ****************************************************9*********************************************
// STEUERUNG: QUERFAHRT
// *************************************************************************************************

IF ( AuftragsdatenStation[wStation].wAuftrag = eStation_Vorabpositionierung ) THEN
  (* Hinweis:
     - Aufruf der Schrittkette
  *)
  Querfahrt[wStation]( Auftragsdaten := AuftragsdatenStation[wStation], wStation := wStation);
  (* Hinweis:
     - Abschluss der Schrittkette
  *)
  IF Querfahrt[wStation].bpDone THEN
    AuftragsdatenStation[wStation] := Querfahrt[wStation].Auftragsdaten;
    Querfahrt[wStation](bpReset := TRUE);
  END_IF
  (* Hinweis:
     - Fehler-Auswertung
  *)
  blFehler[wStation, cWAND_1] := Querfahrt[wStation].bpFehler;
  IF rtlFehler[wStation, cWAND_1].Q THEN
    AutomatikFehlerSetzen(starrShuttleBasisParameter[wStation].stMKs.eaAutomatikkreis, abpFehler);
  END_IF
ELSE
  (* Hinweis:
     - Reset der Schrittkette
  *)
  IF ( Querfahrt[wStation].steplSchritt <> STEP_0_E ) THEN
    Querfahrt[wStation](bpReset := TRUE);
  END_IF
END_IF
END_METHOD

(* ---- ShuttleWandAuftraege.meth.st ---- *)
(* METADATA
{
	"v3Meta": {
		"objectGuid": "a4d875f2-deb1-4181-ad49-6660bcb8c981"
	}
}
*)
METHOD ShuttleWandAuftraege
VAR_INPUT
  wStation : WORD;
  wWand    : WORD;
END_VAR

// ****************************************************9*********************************************
// STEUERUNG: EINTRANSPORT
// *************************************************************************************************

IF ( AuftragsdatenWand[wStation, wWand].wAuftrag = eStation_Eintransport ) THEN
  (* Hinweis:
     - Aufruf der Schrittkette
  *)
  starrShuttleBasisParameter[wStation].bEintransportGewesen[wWand] := FALSE;
  Eintransport[wStation, wWand]( Auftragsdaten := AuftragsdatenWand[wStation, wWand], wStation := wStation, wWand := wWand);
  (* Hinweis:
     - Abschluss der Schrittkette
  *)
  IF Eintransport[wStation, wWand].bpDone THEN
    // Scheibe liegt nur definiert am Stopp-Sensor in Transportrichtung:
    // vorwaerts auf Auslauf mit Auslauf-Stopp, rueckwaerts auf Einlauf mit Einlauf-Stopp
    starrShuttleBasisParameter[wStation].bEintransportGewesen[wWand] :=
         (     NOT starrShuttleBasisParameter[wStation].bRueckwaertsTransportieren[wWand]
           AND ( starrShuttleBasisParameter[wStation].pAuftrag[wWand].stAuftragsOptionen.eGlastransport = eGlastransport_AufAuslauf )
           AND starrShuttleBasisParameter[wStation].stMKs.stStationsAufbau.bSensorAuslaufStopp )
      OR (     starrShuttleBasisParameter[wStation].bRueckwaertsTransportieren[wWand]
           AND ( starrShuttleBasisParameter[wStation].pAuftrag[wWand].stAuftragsOptionen.eGlastransport = eGlastransport_AufEinlauf )
           AND starrShuttleBasisParameter[wStation].stMKs.stStationsAufbau.bSensorEinlaufStopp );
    AuftragsdatenWand[wStation, wWand] := Eintransport[wStation, wWand].Auftragsdaten;
    Eintransport[wStation, wWand](bpReset := TRUE);
  END_IF
  (* Hinweis:
     - Fehler-Auswertung
  *)
  blFehler[wStation, wWand] := Eintransport[wStation, wWand].bpFehler;
  IF rtlFehler[wStation, wWand].Q THEN
    AutomatikFehlerSetzen(starrShuttleBasisParameter[wStation].stMKs.eaAutomatikkreis, abpFehler);
  END_IF
ELSE
  (* Hinweis:
     - Reset der Schrittkette
  *)
  IF ( Eintransport[wStation, wWand].steplSchritt > STEP_0_E ) THEN
    Eintransport[wStation, wWand](bpReset := TRUE);
  END_IF
END_IF

// ****************************************************9*********************************************
// STEUERUNG: AUSTRANSPORT
// *************************************************************************************************

IF ( AuftragsdatenWand[wStation, wWand].wAuftrag = eStation_Austransport ) THEN
  (* Hinweis:
     - Aufruf der Schrittkette
     - bEintransportGewesen bleibt bis zum Ende des Austransports stehen: Die Vorab-Ansteuerung wartet, bis der
       Glastransport den Eintransport beendet hat, und prueft den Merker erst danach (Verbrauch dort)
  *)
  Austransport[wStation, wWand]( Auftragsdaten := AuftragsdatenWand[wStation, wWand], wStation := wStation, wWand := wWand);
  (* Hinweis:
     - Abschluss der Schrittkette
  *)
  IF Austransport[wStation, wWand].bpDone THEN
    starrShuttleBasisParameter[wStation].bEintransportGewesen[wWand] := FALSE;
    AuftragsdatenWand[wStation, wWand] := Austransport[wStation, wWand].Auftragsdaten;
    Austransport[wStation, wWand](bpReset := TRUE);
  END_IF
  (* Hinweis:
     - Fehler-Auswertung
  *)
  blFehler[wStation, wWand] := Austransport[wStation, wWand].bpFehler;
  IF rtlFehler[wStation, wWand].Q THEN
    AutomatikFehlerSetzen(starrShuttleBasisParameter[wStation].stMKs.eaAutomatikkreis, abpFehler);
  END_IF
ELSE
  (* Hinweis:
     - Reset der Schrittkette
  *)
  IF ( Austransport[wStation, wWand].steplSchritt > STEP_0_E ) THEN
    Austransport[wStation, wWand](bpReset := TRUE);
  END_IF
END_IF

// ****************************************************9*********************************************
// STEUERUNG: DURCHTRANSPORT
// *************************************************************************************************

IF ( AuftragsdatenWand[wStation, wWand].wAuftrag = eStation_Durchtransport ) THEN
  (* Hinweis:
     - Aufruf der Schrittkette
  *)
  Durchtransport[wStation, wWand]( Auftragsdaten := AuftragsdatenWand[wStation, wWand], wStation := wStation, wWand := wWand);
  (* Hinweis:
     - Abschluss der Schrittkette
  *)
  IF Durchtransport[wStation, wWand].bpDone THEN
    AuftragsdatenWand[wStation, wWand] := Durchtransport[wStation, wWand].Auftragsdaten;
    Durchtransport[wStation, wWand](bpReset := TRUE);
  END_IF
  (* Hinweis:
     - Fehler-Auswertung
  *)
  blFehler[wStation, wWand] := Durchtransport[wStation, wWand].bpFehler;
  IF rtlFehler[wStation, wWand].Q THEN
    AutomatikFehlerSetzen(starrShuttleBasisParameter[wStation].stMKs.eaAutomatikkreis, abpFehler);
  END_IF
ELSE
  (* Hinweis:
     - Reset der Schrittkette
  *)
  IF ( Durchtransport[wStation, wWand].steplSchritt > STEP_0_E ) THEN
    Durchtransport[wStation, wWand](bpReset := TRUE);
  END_IF
END_IF

// ****************************************************9*********************************************
// STEUERUNG: VORABKOMPONENTEN
// *************************************************************************************************
IF ( VorAbAuftragsDaten[wStation, wWand].wAuftrag = eStation_VorabAuftrag ) THEN
  (* Hinweis:
     - Aufruf der Schrittkette
  *)
  VorabkomponentenAnsteuerung[wStation, wWand]( Auftragsdaten := VorAbAuftragsDaten[wStation, wWand],  wStation := wStation, wWand := wWand);
  (* Hinweis:
     - Abschluss der Schrittkette
  *)
  IF VorabkomponentenAnsteuerung[wStation, wWand].bpDone THEN
    VorAbAuftragsDaten[wStation, wWand] := VorabkomponentenAnsteuerung[wStation, wWand].Auftragsdaten;
    VorabkomponentenAnsteuerung[wStation, wWand](bpReset := TRUE);
  END_IF
  (* Hinweis:
     - Fehler-Auswertung
  *)
  blFehler[wStation, wWand] := VorabkomponentenAnsteuerung[wStation, wWand].bpFehler;
  IF rtlFehler[wStation, wWand].Q THEN
    AutomatikFehlerSetzen(starrShuttleBasisParameter[wStation].stMKs.eaAutomatikkreis, abpFehler);
  END_IF
ELSE
  (* Hinweis:
     - Reset der Schrittkette
  *)
  IF ( VorabkomponentenAnsteuerung[wStation, wWand].steplSchritt > STEP_0_E ) THEN
    VorabkomponentenAnsteuerung[wStation, wWand](bpReset := TRUE);
  END_IF
END_IF

// ****************************************************9*********************************************
// STEUERUNG: RACKSUCHE
// *************************************************************************************************

IF ( AuftragsdatenWand[wStation, wWand].wAuftrag = eStation_RackSuche ) THEN
  (* Hinweis:
     - Aufruf der Schrittkette
  *)
  Racksuche[wStation]( Auftragsdaten := AuftragsdatenWand[wStation, wWand], wStation := wStation );
  (* Hinweis:
     - Abschluss der Schrittkette
  *)
  IF Racksuche[wStation].bpDone THEN
    AuftragsdatenWand[wStation, wWand] := Racksuche[wStation].Auftragsdaten;
    Racksuche[wStation](bpReset := TRUE);
  END_IF
  (* Hinweis:
     - Fehler-Auswertung
  *)
  blFehler[wStation, cWAND_1] := Racksuche[wStation].bpFehler;
  IF rtlFehler[wStation, cWAND_1].Q THEN
    AutomatikFehlerSetzen(starrShuttleBasisParameter[wStation].stMKs.eaAutomatikkreis, abpFehler);
  END_IF
ELSE
  (* Hinweis:
     - Reset der Schrittkette
  *)
  IF ( Racksuche[wStation].steplSchritt <> STEP_0_E ) THEN
    Racksuche[wStation](bpReset := TRUE);
  END_IF
END_IF
END_METHOD

(* ---- Slave_Transfershuttle.meth.st ---- *)
(* METADATA
{
	"v3Meta": {
		"objectGuid": "0f9ee576-0110-44f2-822b-96aae40b0d13"
	}
}
*)
METHOD INTERNAL Slave_Transfershuttle
VAR_INPUT
  wStation : WORD;
END_VAR

// ****************************************************9*********************************************
// STEUERUNG: TRANSPORTKOPPLUNG
// *************************************************************************************************

IF ( AuftragsdatenTransfershuttle[wStation].wAuftrag = eStation_Transportkopplung ) THEN
  (* Hinweis:
     - Aufruf der Schrittkette
  *)
  TS_Transportkopplung[wStation]( Auftragsdaten := AuftragsdatenTransfershuttle[wStation], wStation := wStation );
  (* Hinweis:
     - Fehler-Auswertung
  *)
  blFehlerTS[wStation] := TS_Transportkopplung[wStation].bpFehler;
  IF rtlFehlerTS[wStation].Q THEN
    CASE AuftragsdatenTransfershuttle[wStation - 1].wAuftrag OF
      eStation_Eintransport:
        IF ( ( awlGlasSender[wStation - 1] >= cERSTES_INPUTSHUTTLE )
             AND ( awlGlasSender[wStation - 1] <= cLETZTES_INPUTSHUTTLE ) )
        THEN
          AutomatikFehlerTransfershuttleSetzen(starrTransferShuttleBasisParameter[wStation].stMKs.eaAutomatikkreis, abpFehler, cSPEICHER_EINLAUFSEITE);
        ELSIF ( ( awlGlasSender[wStation - 1] >= cERSTES_OUTPUTSHUTTLE )
                AND ( awlGlasSender[wStation - 1] <= cLETZTES_OUTPUTSHUTTLE ) )
        THEN
          AutomatikFehlerTransfershuttleSetzen(starrTransferShuttleBasisParameter[wStation].stMKs.eaAutomatikkreis, abpFehler, cSPEICHER_AUSLAUFSEITE);
        ELSE
          AutomatikFehlerSetzen(starrTransferShuttleBasisParameter[wStation].stMKs.eaAutomatikkreis, abpFehler);
        END_IF
      eStation_Austransport:
        IF ( ( awlGlasSender[wStation - 1] >= cERSTES_OUTPUTSHUTTLE )
             AND ( awlGlasSender[wStation - 1] <= cLETZTES_OUTPUTSHUTTLE ) )
        THEN
          AutomatikFehlerTransfershuttleSetzen(starrTransferShuttleBasisParameter[wStation].stMKs.eaAutomatikkreis, abpFehler, cSPEICHER_EINLAUFSEITE);
        ELSIF ( ( awlGlasSender[wStation - 1] >= cERSTES_INPUTSHUTTLE )
                AND ( awlGlasSender[wStation - 1] <= cLETZTES_INPUTSHUTTLE ) )
        THEN
          AutomatikFehlerTransfershuttleSetzen(starrTransferShuttleBasisParameter[wStation].stMKs.eaAutomatikkreis, abpFehler, cSPEICHER_AUSLAUFSEITE);
        ELSE
          AutomatikFehlerSetzen(starrTransferShuttleBasisParameter[wStation].stMKs.eaAutomatikkreis, abpFehler);
        END_IF
      eStation_Vortransport:
        AutomatikFehlerSetzen(starrTransferShuttleBasisParameter[wStation].stMKs.eaAutomatikkreis, abpFehler);
      ELSE
        IF atonlWarteAufMasterAuftrag[wStation].Q THEN
          AutomatikFehlerSetzen(starrTransferShuttleBasisParameter[wStation].stMKs.eaAutomatikkreis, abpFehler);
        END_IF
    END_CASE
  END_IF
ELSE
  (* Hinweis:
     - Reset der Schrittkette
  *)
  IF ( TS_Transportkopplung[wStation].steplSchritt <> STEP_0_E ) THEN
    TS_Transportkopplung[wStation](bpReset := TRUE);
  END_IF
END_IF

// ****************************************************9*********************************************
// STEUERUNG: QUERFAHRT
// *************************************************************************************************

IF ( AuftragsdatenTransfershuttle[wStation].wAuftrag = eStation_Vorabpositionierung ) THEN
  (* Hinweis:
     - Aufruf der Schrittkette
  *)
  TS_Querfahrt[wStation]( Auftragsdaten := AuftragsdatenTransfershuttle[wStation], wStation := wStation );
  (* Hinweis:
     - Abschluss der Schrittkette
  *)
  IF TS_Querfahrt[wStation].bpDone THEN
    AuftragsdatenTransfershuttle[wStation] := Querfahrt[wStation].Auftragsdaten;
    TS_Querfahrt[wStation](bpReset := TRUE);
  END_IF
  (* Hinweis:
     - Fehler-Auswertung
  *)
  blFehlerTS[wStation] := TS_Querfahrt[wStation].bpFehler;
  IF rtlFehlerTS[wStation].Q THEN
    AutomatikFehlerSetzen(starrTransferShuttleBasisParameter[wStation].stMKs.eaAutomatikkreis, abpFehler);
  END_IF
ELSE
  (* Hinweis:
     - Reset der Schrittkette
  *)
  IF ( TS_Querfahrt[wStation].steplSchritt <> STEP_0_E ) THEN
    TS_Querfahrt[wStation](bpReset := TRUE);
  END_IF
END_IF
END_METHOD

(* ---- Verfahrfreigabe.act.st ---- *)
(* METADATA
{
	"v3Meta": {
		"objectGuid": "c5ed0ecf-290a-4d28-a44b-5709f6fc01b5"
	}
}
*)
ACTION Verfahrfreigabe
//-------------------------------------------------------------------------------------------------
// BAUSTEIN: VERFAHRFREIGABE SHUTTLE
//-------------------------------------------------------------------------------------------------
(* Hinweis:
   - bpShuttleAnhalten wird generisch aus starrShuttleBasisParameter[...].stMKs.astShuttleAnhaltenQuellen gebildet.
   - Pro Shuttle werden alle aktiven Eintraege per OR verknuepft.
   - Keine festen Stations- oder Shuttle-Nummern im Code.
   - Parametrierung erfolgt ausschliesslich in MK_Shuttle.
   - getBasis() loest Station / Shuttle / Transfershuttle einheitlich auf.
*)
FOR wlIndex := cERSTES_SHUTTLE TO cLETZTES_SHUTTLE DO

  aShuttle[wlIndex].bpShuttleAnhalten := FALSE;

  FOR wlIndexQuelle := 1 TO cMAX_SHUTTLE_ANHALTEN_QUELLEN DO

    IF starrShuttleBasisParameter[wlIndex].stMKs.astShuttleAnhaltenQuellen[wlIndexQuelle].bAktiv THEN

      Basis REF= getBasis(starrShuttleBasisParameter[wlIndex].stMKs.astShuttleAnhaltenQuellen[wlIndexQuelle].wQuellenNummer);

      // Hinweis: Quelle ist in dieser Konfiguration nicht vorhanden => ueberspringen
      IF __ISVALIDREF( Basis ) THEN

        CASE starrShuttleBasisParameter[wlIndex].stMKs.astShuttleAnhaltenQuellen[wlIndexQuelle].eSensorTyp OF

          eAuslaufsensor:
            IF Basis.OutGlasTransport[starrShuttleBasisParameter[wlIndex].stMKs.astShuttleAnhaltenQuellen[wlIndexQuelle].wWand].bScheibeFaehrtUeberAuslauf THEN
              aShuttle[wlIndex].bpShuttleAnhalten := TRUE;
            END_IF

          eEinlaufsensor:
            IF Basis.OutGlasTransport[starrShuttleBasisParameter[wlIndex].stMKs.astShuttleAnhaltenQuellen[wlIndexQuelle].wWand].bScheibeFaehrtUeberEinlauf THEN
              aShuttle[wlIndex].bpShuttleAnhalten := TRUE;
            END_IF

        END_CASE

      END_IF

    END_IF

  END_FOR

END_FOR

// ---------------------------------------------------------------------------------------
//  VERFAHRLOGIK - RESET DER POSITIONIERUNG NACH ABBRUCH
//
//  Hinweis:
//  - Zurueck des Auftrags  "cSHUTTLE_VORABPOSITIONIERUNG" wenn dieser aktiv gewesen ist
// ---------------------------------------------------------------------------------------
FOR wlIndex := cERSTES_SHUTTLE TO cLETZTES_SHUTTLE DO
  IF  ( starrShuttleBasisParameter[wlIndex].bPositionierAuftragZuruecksetzen ) THEN
    IF ( AuftragsdatenStation[wlIndex].wAuftrag = eStation_Vorabpositionierung ) THEN
      starrShuttleBasisParameter[wlIndex].bQuittungPositionierungZurueckgesetzt := TRUE;
      AuftragsdatenStation[wlIndex].wAuftrag := eStation_Kein_Auftrag;
    END_IF
  END_IF
END_FOR

// ---------------------------------------------------------------------------------------
//  VERFAHRLOGIK TRANSFERSHUTTLE - RESET DER POSITIONIERUNG NACH ABBRUCH
//
//  Hinweis:
//  - Zurueck des Auftrags  "cSHUTTLE_VORABPOSITIONIERUNG" wenn dieser aktiv gewesen ist
// ---------------------------------------------------------------------------------------
FOR wlIndex := cERSTES_TRANSFERSHUTTLE TO cLETZTES_TRANSFERSHUTTLE DO
  IF  ( starrTransfershuttleBasisParameter[wlIndex].bPositionierAuftragZuruecksetzen ) THEN
    IF ( AuftragsdatenTransfershuttle[wlIndex].wAuftrag = eStation_Vorabpositionierung ) THEN
      starrTransfershuttleBasisParameter[wlIndex].bQuittungPositionierungZurueckgesetzt := TRUE;
      AuftragsdatenTransfershuttle[wlIndex].wAuftrag := eStation_Kein_Auftrag;
    END_IF
  END_IF
END_FOR
END_ACTION

(* ---- Visu.act.st ---- *)
(* METADATA
{
	"v3Meta": {
		"objectGuid": "1e9e5d8c-b3c6-4e22-b591-305900ce7097"
	}
}
*)
ACTION Visu
//-------------------------------------------------------------------------------------------------
// Daten in das VisoArray kopieren
//-------------------------------------------------------------------------------------------------

FOR wlIndex := cERSTES_SHUTTLE TO cLETZTES_SHUTTLE DO
  VisuAuftragsdaten[wlIndex].eStation := TO_WORD(AuftragsdatenStation[wlIndex].wAuftrag);
  FOR wlIndexWand := cWAND_1 TO cANZAHL_WAENDE DO
    VisuAuftragsdaten[wlIndex].eWand[wlIndexWand] := TO_WORD(AuftragsdatenWand[wlIndex, wlIndexWand].wAuftrag);
  END_FOR
END_FOR

FOR wlIndex := cERSTES_TRANSFERSHUTTLE TO cLETZTES_TRANSFERSHUTTLE DO
  VisuAuftragsdaten[wlIndex].eStation := TO_WORD(AuftragsdatenTransfershuttle[wlIndex].wAuftrag);
END_FOR
END_ACTION
